(* IEC 61131-3 sources: Lasal-MCP/examples/SampleSource/LASALScreenAdvancedSolution/LASALScreenAdvancedSolution/LASALScreenAdvacnedSolution/Stations/MachineControl/MachineControl/Network/STDCommunicationToHMI, 1 file *)

(* ---- ONE_STDCommunicationToHMI_Table.st ---- *)
#define OBJECTS_CONFIG

#include "..\..\Class\_AlarmX0Para\_AlarmX0Para.h"
#include "..\..\Class\DataManager\DataManager.h"
//Define part of class DataManagerFIFO
#define MEMORY_Mark_DataMngFiFo    8
#include <.\lsl_st_mt.h>
#include "..\..\Class\TCPCommunication\TCPCommunication.h"
#include "..\..\Class\TCPCommunication\SalamanderDelay.h"

FUNCTION GLOBAL TAB ONE_STDCommunicationToHMI
-1$UINT, 0$UINT,
1$UINT, 0$UINT,

14$UDINT,
TO_UDINT(800276940), "_AlarmX0Para", 0$UINT, 11$UINT, 1$UINT,
TO_UDINT(3900434542), "_CheckOnlineStatus", 1$UINT, 4$UINT, 1$UINT,
TO_UDINT(916194998), "_CheckSum", 1$UINT, 0$UINT, 1$UINT,
TO_UDINT(794617671), "CriticalSection", 0$UINT, 4$UINT, 10$UINT,
TO_UDINT(4008337867), "DataManager", 1$UINT, 1$UINT, 1$UINT,
TO_UDINT(2873804345), "DataManagerFIFO", 1$UINT, 0$UINT, 10$UINT,
TO_UDINT(2393054465), "DataManagerPriority", 1$UINT, 0$UINT, 1$UINT,
TO_UDINT(2602835227), "GetTaskHandle", 0$UINT, 2$UINT, 1$UINT,
TO_UDINT(2225119864), "MerkerEx", 1$UINT, 22$UINT, 2$UINT,
TO_UDINT(3534980377), "RamRingBuffer", 1$UINT, 1$UINT, 1$UINT,
TO_UDINT(1850111279), "String", 1$UINT, 11$UINT, 1$UINT,
TO_UDINT(2898603620), "StringInternal", 1$UINT, 85$UINT, 0$UINT,
TO_UDINT(3704218787), "TCPCommunication", 1$UINT, 17$UINT, 1$UINT,
TO_UDINT(3232495061), "VirtualBaseInit", 1$UINT, 3$UINT, 0$UINT,

_NO_ATTR, TO_UDINT(2051489927), "ALARMCOMMUNICATION",

_NO_ATTR, TO_UDINT(2314772430), "CHECKONLINESTATUS1",

1$UINT, TO_UDINT(1168159097), "STDTCPCOMMUNICATIONTOHMI\CHECKSUM",

1$UINT, TO_UDINT(2590012171), "STDDATAMANAGERTOHMI\DATAMANAGERPRIORITY\DATAMANAGERFIFO_PRIO0\SECTION",
1$UINT, TO_UDINT(2367383368), "STDDATAMANAGERTOHMI\DATAMANAGERPRIORITY\DATAMANAGERFIFO_PRIO1\SECTION",
1$UINT, TO_UDINT(3029752717), "STDDATAMANAGERTOHMI\DATAMANAGERPRIORITY\DATAMANAGERFIFO_PRIO2\SECTION",
1$UINT, TO_UDINT(2750238670), "STDDATAMANAGERTOHMI\DATAMANAGERPRIORITY\DATAMANAGERFIFO_PRIO3\SECTION",
1$UINT, TO_UDINT(3347849735), "STDDATAMANAGERTOHMI\DATAMANAGERPRIORITY\DATAMANAGERFIFO_PRIO4\SECTION",
1$UINT, TO_UDINT(3505862212), "STDDATAMANAGERTOHMI\DATAMANAGERPRIORITY\DATAMANAGERFIFO_PRIO5\SECTION",
1$UINT, TO_UDINT(3917089409), "STDDATAMANAGERTOHMI\DATAMANAGERPRIORITY\DATAMANAGERFIFO_PRIO6\SECTION",
1$UINT, TO_UDINT(4261486274), "STDDATAMANAGERTOHMI\DATAMANAGERPRIORITY\DATAMANAGERFIFO_PRIO7\SECTION",
1$UINT, TO_UDINT(565760275), "STDDATAMANAGERTOHMI\DATAMANAGERPRIORITY\DATAMANAGERFIFO_PRIO8\SECTION",
1$UINT, TO_UDINT(918799696), "STDDATAMANAGERTOHMI\DATAMANAGERPRIORITY\DATAMANAGERFIFO_PRIO9\SECTION",

_NO_ATTR, TO_UDINT(4280838709), "STDDATAMANAGERTOHMI",

1$UINT, TO_UDINT(3236025859), "STDDATAMANAGERTOHMI\DATAMANAGERPRIORITY\DATAMANAGERFIFO_PRIO0",
1$UINT, TO_UDINT(3085362837), "STDDATAMANAGERTOHMI\DATAMANAGERPRIORITY\DATAMANAGERFIFO_PRIO1",
1$UINT, TO_UDINT(787461935), "STDDATAMANAGERTOHMI\DATAMANAGERPRIORITY\DATAMANAGERFIFO_PRIO2",
1$UINT, TO_UDINT(1508411321), "STDDATAMANAGERTOHMI\DATAMANAGERPRIORITY\DATAMANAGERFIFO_PRIO3",
1$UINT, TO_UDINT(3347845658), "STDDATAMANAGERTOHMI\DATAMANAGERPRIORITY\DATAMANAGERFIFO_PRIO4",
1$UINT, TO_UDINT(2961908364), "STDDATAMANAGERTOHMI\DATAMANAGERPRIORITY\DATAMANAGERFIFO_PRIO5",
1$UINT, TO_UDINT(696415030), "STDDATAMANAGERTOHMI\DATAMANAGERPRIORITY\DATAMANAGERFIFO_PRIO6",
1$UINT, TO_UDINT(1585791904), "STDDATAMANAGERTOHMI\DATAMANAGERPRIORITY\DATAMANAGERFIFO_PRIO7",
1$UINT, TO_UDINT(3459931697), "STDDATAMANAGERTOHMI\DATAMANAGERPRIORITY\DATAMANAGERFIFO_PRIO8",
1$UINT, TO_UDINT(3107810983), "STDDATAMANAGERTOHMI\DATAMANAGERPRIORITY\DATAMANAGERFIFO_PRIO9",

1$UINT, TO_UDINT(3371365168), "STDDATAMANAGERTOHMI\DATAMANAGERPRIORITY",

1$UINT, TO_UDINT(1559645213), "STDDATAMANAGERTOHMI\DATAMNGGETTASKHANDLE1",

1$UINT, TO_UDINT(746981269), "STDTCPCOMMUNICATIONTOHMI\RAMRINGMERKEREX",
1$UINT, TO_UDINT(1992695623), "STDTCPCOMMUNICATIONTOHMI\THREADNAME\MERKEREX0",

1$UINT, TO_UDINT(3210803935), "STDTCPCOMMUNICATIONTOHMI\RAMRINGBUFFER",

1$UINT, TO_UDINT(1839612986), "STDTCPCOMMUNICATIONTOHMI\THREADNAME",

_NO_ATTR, TO_UDINT(1352039343), "STDTCPCOMMUNICATIONTOHMI",

//Internal connections
0$UDINT,
27$UDINT,
TO_UDINT(13), "DataMngGetTaskHandle1", TO_UDINT(25),
TO_UDINT(13), "DataManagerPriority", TO_UDINT(24),
TO_UDINT(14), "Section", TO_UDINT(3),
TO_UDINT(15), "Section", TO_UDINT(4),
TO_UDINT(16), "Section", TO_UDINT(5),
TO_UDINT(17), "Section", TO_UDINT(6),
TO_UDINT(18), "Section", TO_UDINT(7),
TO_UDINT(19), "Section", TO_UDINT(8),
TO_UDINT(20), "Section", TO_UDINT(9),
TO_UDINT(21), "Section", TO_UDINT(10),
TO_UDINT(22), "Section", TO_UDINT(11),
TO_UDINT(23), "Section", TO_UDINT(12),
TO_UDINT(24), "DataManagerFiFo_Prio0", TO_UDINT(14),
TO_UDINT(24), "DataManagerFiFo_Prio1", TO_UDINT(15),
TO_UDINT(24), "DataManagerFiFo_Prio2", TO_UDINT(16),
TO_UDINT(24), "DataManagerFiFo_Prio3", TO_UDINT(17),
TO_UDINT(24), "DataManagerFiFo_Prio4", TO_UDINT(18),
TO_UDINT(24), "DataManagerFiFo_Prio5", TO_UDINT(19),
TO_UDINT(24), "DataManagerFiFo_Prio6", TO_UDINT(20),
TO_UDINT(24), "DataManagerFiFo_Prio7", TO_UDINT(21),
TO_UDINT(24), "DataManagerFiFo_Prio8", TO_UDINT(22),
TO_UDINT(24), "DataManagerFiFo_Prio9", TO_UDINT(23),
TO_UDINT(29), "MerkerEx0", TO_UDINT(27),
TO_UDINT(30), "RamRingBuffer", TO_UDINT(28),
TO_UDINT(30), "RamRingMerkerEx", TO_UDINT(26),
TO_UDINT(30), "CheckSum", TO_UDINT(2),
TO_UDINT(30), "ThreadName", TO_UDINT(29),
0$UDINT,
6$UDINT,
TO_UDINT(1), "toTCPComm", TO_UDINT(30), "ClassSvr",
TO_UDINT(1), "AlarmCommunication", TO_UDINT(0), "ClassSvr",
TO_UDINT(13), "coTCPCommunication", TO_UDINT(30), "ClassSvr",
TO_UDINT(28), "Data", TO_UDINT(26), "m_udLength",
TO_UDINT(29), "DataBuffer", TO_UDINT(27), "m_udLength",
TO_UDINT(30), "coDataMng", TO_UDINT(13), "ClassSvr",

//Initialization values
0$UDINT,
12$UDINT,
TO_UDINT(0), "Config", TO_UDINT(0),//|STDCommunicationToHMI.AlarmCommunication.Config;
TO_UDINT(1), "DelayTime", TO_UDINT(20000),//|STDCommunicationToHMI.CheckOnlineStatus1.DelayTime;
TO_UDINT(13), "AcceptOfflineJobs", TO_UDINT(1),//|STDCommunicationToHMI.STDDataManagerToHMI.AcceptOfflineJobs;
TO_UDINT(26), "ThreadSafe", TO_UDINT(0),//|STDCommunicationToHMI.STDTCPCommunicationToHMI\RamRingMerkerEx.ThreadSafe;
TO_UDINT(27), "ThreadSafe", TO_UDINT(0),//|STDCommunicationToHMI.ThreadName\STDTCPCommunicationToHMI\MerkerEx0.ThreadSafe;
TO_UDINT(29), "SingleRealloc", TO_UDINT(1),//|STDCommunicationToHMI.STDTCPCommunicationToHMI\ThreadName.SingleRealloc;
TO_UDINT(30), "ComPort", TO_UDINT(500),//|STDCommunicationToHMI.STDTCPCommunicationToHMI.ComPort;
TO_UDINT(30), "LogEnable", TO_UDINT(0),//|STDCommunicationToHMI.STDTCPCommunicationToHMI.LogEnable;
TO_UDINT(30), "DeactivateCom", TO_UDINT(0),//|STDCommunicationToHMI.STDTCPCommunicationToHMI.DeactivateCom;
TO_UDINT(30), "coLogFilter", TO_UDINT(0),//|STDCommunicationToHMI.STDTCPCommunicationToHMI.coLogFilter;
TO_UDINT(30), "SizeOfComBuffers", TO_UDINT(2MB),//|STDCommunicationToHMI.STDTCPCommunicationToHMI.SizeOfComBuffers;
TO_UDINT(30), "SizeOfComBufferRecv", TO_UDINT(2MB),//|STDCommunicationToHMI.STDTCPCommunicationToHMI.SizeOfComBufferRecv;

//Symbolic initialization values
0$UDINT,
0$UDINT,

//Initialization of string values
0$UDINT,
0$UDINT,

//Configuration of tasks (RealTime, Cyclic, Background)
0$UDINT,
1$UDINT,
TO_UDINT(25), (1000)$UDINT, 4194303$DINT, 	//STDDATAMANAGERTOHMI\DATAMNGGETTASKHANDLE1

0$UDINT,
3$UDINT,
TO_UDINT(1), (50)$UDINT, 4194303$DINT, 	//CHECKONLINESTATUS1
TO_UDINT(25), (1000)$UDINT, 4194303$DINT, 	//STDDATAMANAGERTOHMI\DATAMNGGETTASKHANDLE1
TO_UDINT(30), (100)$UDINT, 4194303$DINT, 	//STDTCPCOMMUNICATIONTOHMI

0$UDINT,
1$UDINT,
TO_UDINT(25), (1000)$UDINT, 4194303$DINT, 	//STDDATAMANAGERTOHMI\DATAMNGGETTASKHANDLE1

//External connections
0$UDINT,
0$UDINT,

//Magic internal connections
0$UDINT,
0$UDINT,

//Configuration of timeslots of tasks (RealTime, Cyclic)
#ifdef __LSLLDR_TIMESLOTS__
0$UDINT,
0$UDINT,

0$UDINT,
0$UDINT,

#endif //__LSLLDR_TIMESLOTS__

//MultiMaster connections
#ifdef __LSLLDR_MULTIMASTER__
0$UDINT,
0$UDINT,
#endif //__LSLLDR_MULTIMASTER__

//Configuration for task ID (RealTime, CyclicTime)
#ifdef __LSLLDR_TASKID__
"\\\\TASKS2  "
0$UDINT,
1$UDINT,
(0)$UDINT, 	//STDDATAMANAGERTOHMI\DATAMNGGETTASKHANDLE1

0$UDINT,
3$UDINT,
(0)$UDINT, 	//CHECKONLINESTATUS1
(0)$UDINT, 	//STDDATAMANAGERTOHMI\DATAMNGGETTASKHANDLE1
(0)$UDINT, 	//STDTCPCOMMUNICATIONTOHMI

0$UDINT,
1$UDINT,
(0)$UDINT, 	//STDDATAMANAGERTOHMI\DATAMNGGETTASKHANDLE1

#endif //__LSLLDR_TASKID__

END_FUNCTION
